(* IEC 61131-3 sources: st-analyze/src, 1 file *)

(* ---- qqqqqqqqqqqqqqq.st ---- *)
TYPE
	City: STRUCT
	 cityId: INT;
	 region: Region;
	 dtTimeNow: DATE_AND_TIME := DT#2021 - 10 - 19 - 13: 53: 00;
   END_STRUCT
END_TYPE
